Staubli VAL3: getAngIOSize.pgx

public program getAngIOSize(num& x_nSize)
  local num l_nSize
begin
  switch rs:sBusUsing
    case "MODBUS"
      l_nSize=size(_aInModbus)
    break
    case "PROFINET"
      l_nSize=size(_aInProfinet)
    break
    case "PROFIBUS"
      l_nSize=size(_aInProfibus)
    break
    case "ETHERCAT"
      l_nSize=size(_aInEthercat)
    break
    case "ETHERNET"
      l_nSize=size(_aInEthernet)
    break
  endSwitch
  x_nSize=l_nSize
end
